FUNCTION_BLOCK FB_mF_Test EXTENDS TcUnit.FB_TestSuite

valueShouldChangeWhenInputChangesAfter1Cycle();

METHOD valueShouldChangeWhenInputChangesAfter1Cycle
VAR
	mF : FB_mF;
	uTest : ARRAY[1..15] OF LREAL;
END_VAR

TEST('valueShouldChangeWhenInputChangesAfter1Cycle');
	mF.setParams(
		activateObserver := FALSE);
	uTest[1] := 50;
	mF.Step(
			u := uTest,
			yMeas := 2);
			
	// After 1 cycle passed, call the model again
	mF.Step(
			u := uTest,
			yMeas := 2);
			
	AssertEquals_BOOL(Expected :=  TRUE, Actual := mF.y[1] <> 0, Message := 'Deviation not zero when current flow is zero');	
TEST_FINISHED();
END_METHOD

END_FUNCTION_BLOCK

(* stored: Version 1.1.0.1, ProductVersion 3.1.4024.9
   POU FB_mF_Test: Id {708b8679-5820-4e1a-b12f-14fefcaf4b3f}, SpecialFunc None
   Method valueShouldChangeWhenInputChangesAfter1Cycle: Id {b5b7ab4d-439e-4b12-a44f-3e31034fb820} *)
